Fanuc KAREL source: kf00087.KL

-- PROVISIONAL review KL for V1013-1; original PC SHA256 3b7f4306b4fdd5ec90424de67af1a70051a7fb9f3e18da821c896b04c0185ce3
-- Incomplete behavior may be omitted. Consult companion uncertainty JSON. Do not deploy.
PROGRAM KF00087
%NOLOCKGROUP
BEGIN
  -- UNRESOLVED_PC offsets 5-28; opcodes 27,22,1C,31,4A
  -- UNRESOLVED_PC offsets 33-37; opcodes 7F
END KF00087
